FUNCTION_BLOCK MGE_Generico (* Multimedidor PM5300 - HidrycoLib *)
  (* Standard: 61499-2 *)
  (* Version 1.5, 15/10/2026, Hidryco, Hidryco, 1.5: tags de valores do IThis com prefixo STS_ (STS_TENSAO_*, STS_CORRENTE_*, STS_POTENCIA_*, STS_FATOR_POTENCIAL_TOTAL, STS_FREQUENCIA). 1.4: corrente A, B e C baixa (STP_CORRENTE_L, 3 alarmes, retardo STP_TEMPO_CORRENTE). 1.3: so as grandezas, ajustes e alarmes da especificacao do cliente (tensoes AB/BC/CA/AN/BN/CN, correntes A/B/C, potencias ativa e reativa A/B/C/total, frequencia, FP e aparente total; alarmes de comunicacao, FP baixo, tensao FF/FN alta/baixa, corrente A/B/C alta e frequencia alta/baixa). Referencia 0 = alarme desligado; um tempo de retardo por grupo. Os grupos de symlink continuam assinando tudo o que o PM53xxMbtcp publica, mas so as grandezas da especificacao entram na logica. 1.2: alarmes conforme a lista do cliente - falta de fase, tensao FF alta/baixa, tensao FN alta/baixa, corrente A/B/C alta, FP baixo, frequencia alta/baixa e falha de comunicacao (sai a corrente L). 1.1: Frequency do PM53xxMbtcp e VTQLINT: stsFrequencia passa para o grupo das energias (VTQLINT). 1.0: multimedidor PowerLogic PM5300 lido pelo HW CAT SE.FieldDevice.PM53xxMbtcp. Os symlinks do HW CAT (VTQREAL/VTQLINT) apontam para ${PATH}stsTensaoAB ... ${PATH}stsEnergiaAparente e ${PATH}stsComunicacaoOK/stsConexao/stsConexaoInt. Falta de fase, tensao H/L e corrente H/L ajustaveis na IHM (memorizados ate o reset). Tags do IThis com os nomes do CAT MGE antigo. *)
  PACKAGE Hidryco.HidrycoLib;
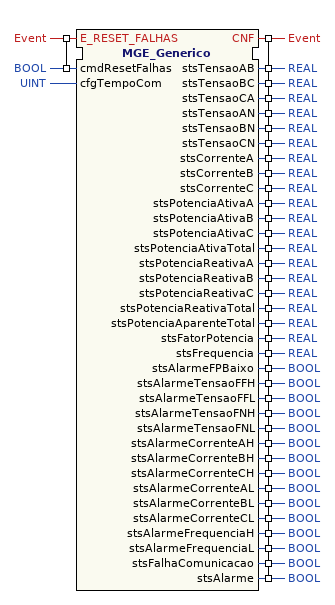
  EVENT_INPUT
    E_RESET_FALHAS WITH cmdResetFalhas; (* Reset pelo processo com cmdResetFalhas = TRUE *)
  END_EVENT
  EVENT_OUTPUT
    CNF WITH stsTensaoAB, stsTensaoBC, stsTensaoCA, stsTensaoAN, stsTensaoBN, stsTensaoCN, stsCorrenteA, stsCorrenteB, stsCorrenteC, stsPotenciaAtivaA, stsPotenciaAtivaB, stsPotenciaAtivaC, stsPotenciaAtivaTotal, stsPotenciaReativaA, stsPotenciaReativaB, stsPotenciaReativaC, stsPotenciaReativaTotal, stsPotenciaAparenteTotal, stsFatorPotencia, stsFrequencia, stsAlarmeFPBaixo, stsAlarmeTensaoFFH, stsAlarmeTensaoFFL, stsAlarmeTensaoFNH, stsAlarmeTensaoFNL, stsAlarmeCorrenteAH, stsAlarmeCorrenteBH, stsAlarmeCorrenteCH, stsAlarmeCorrenteAL, stsAlarmeCorrenteBL, stsAlarmeCorrenteCL, stsAlarmeFrequenciaH, stsAlarmeFrequenciaL, stsFalhaComunicacao, stsAlarme; (* Valores e alarmes (so na mudanca) *)
  END_EVENT
  VAR_INPUT
    cmdResetFalhas : BOOL; (* TRUE = reset (com o evento E_RESET_FALHAS) *)
    cfgTempoCom : UINT := 5; (* Tempo (s) sem comunicacao com o medidor para confirmar a falha *)
  END_VAR
  VAR_OUTPUT
    stsTensaoAB : REAL; (* Tensao A-B (V) *)
    stsTensaoBC : REAL; (* Tensao B-C (V) *)
    stsTensaoCA : REAL; (* Tensao C-A (V) *)
    stsTensaoAN : REAL; (* Tensao A-N (V) *)
    stsTensaoBN : REAL; (* Tensao B-N (V) *)
    stsTensaoCN : REAL; (* Tensao C-N (V) *)
    stsCorrenteA : REAL; (* Corrente fase A (A) *)
    stsCorrenteB : REAL; (* Corrente fase B (A) *)
    stsCorrenteC : REAL; (* Corrente fase C (A) *)
    stsPotenciaAtivaA : REAL; (* Potencia ativa fase A (kW) *)
    stsPotenciaAtivaB : REAL; (* Potencia ativa fase B (kW) *)
    stsPotenciaAtivaC : REAL; (* Potencia ativa fase C (kW) *)
    stsPotenciaAtivaTotal : REAL; (* Potencia ativa total (kW) *)
    stsPotenciaReativaA : REAL; (* Potencia reativa fase A (kVAr) *)
    stsPotenciaReativaB : REAL; (* Potencia reativa fase B (kVAr) *)
    stsPotenciaReativaC : REAL; (* Potencia reativa fase C (kVAr) *)
    stsPotenciaReativaTotal : REAL; (* Potencia reativa total (kVAr) *)
    stsPotenciaAparenteTotal : REAL; (* Potencia aparente total (kVA) *)
    stsFatorPotencia : REAL; (* Fator de potencia total *)
    stsFrequencia : REAL; (* Frequencia (Hz) *)
    stsAlarmeFPBaixo : BOOL; (* Fator de potência baixo (memorizado ate o reconhecimento) *)
    stsAlarmeTensaoFFH : BOOL; (* Tensão entre fases alta (memorizado ate o reconhecimento) *)
    stsAlarmeTensaoFFL : BOOL; (* Tensão entre fases baixa (memorizado ate o reconhecimento) *)
    stsAlarmeTensaoFNH : BOOL; (* Tensão fase-neutro alta (memorizado ate o reconhecimento) *)
    stsAlarmeTensaoFNL : BOOL; (* Tensão fase-neutro baixa (memorizado ate o reconhecimento) *)
    stsAlarmeCorrenteAH : BOOL; (* Corrente fase A alta (memorizado ate o reconhecimento) *)
    stsAlarmeCorrenteBH : BOOL; (* Corrente fase B alta (memorizado ate o reconhecimento) *)
    stsAlarmeCorrenteCH : BOOL; (* Corrente fase C alta (memorizado ate o reconhecimento) *)
    stsAlarmeCorrenteAL : BOOL; (* Corrente fase A baixa (memorizado ate o reconhecimento) *)
    stsAlarmeCorrenteBL : BOOL; (* Corrente fase B baixa (memorizado ate o reconhecimento) *)
    stsAlarmeCorrenteCL : BOOL; (* Corrente fase C baixa (memorizado ate o reconhecimento) *)
    stsAlarmeFrequenciaH : BOOL; (* Frequência alta (memorizado ate o reconhecimento) *)
    stsAlarmeFrequenciaL : BOOL; (* Frequência baixa (memorizado ate o reconhecimento) *)
    stsFalhaComunicacao : BOOL; (* Falha de comunicacao com o medidor *)
    stsAlarme : BOOL; (* Algum alarme do medidor *)
  END_VAR
  FBS
    IThis : MGE_Generico_HMI(QI := TRUE);
    plcStart1 : plcStart(Prio := 10);
    Logica : basicMGEGenerico;
    Tick : E_CYCLE(DT := T#1s);
    Tensoes : SYMLINKMULTIVARDST_2295B2715D3FE1C95(NAME1 := '$${PATH}stsTensaoAB', NAME2 := '$${PATH}stsTensaoBC', NAME3 := '$${PATH}stsTensaoCA', NAME4 := '$${PATH}stsTensaoMediaLL', NAME5 := '$${PATH}stsTensaoAN', NAME6 := '$${PATH}stsTensaoBN', NAME7 := '$${PATH}stsTensaoCN', NAME8 := '$${PATH}stsTensaoMediaLN', NAME9 := '$${PATH}stsDesequilibrioTensao', QI := TRUE); {SET_ATTRIBUTE(Configuration.GenericFBType.InterfaceParams, Runtime.System#I:=9;VALUE${I$}:VTQREAL,VTQREAL,VTQREAL,VTQREAL,VTQREAL,VTQREAL,VTQREAL,VTQREAL,VTQREAL)}
    Correntes : SYMLINKMULTIVARDST_858FA8D101163416(NAME1 := '$${PATH}stsCorrenteA', NAME2 := '$${PATH}stsCorrenteB', NAME3 := '$${PATH}stsCorrenteC', NAME4 := '$${PATH}stsCorrenteMedia', QI := TRUE); {SET_ATTRIBUTE(Configuration.GenericFBType.InterfaceParams, Runtime.System#I:=4;VALUE${I$}:VTQREAL,VTQREAL,VTQREAL,VTQREAL)}
    Potencias : SYMLINKMULTIVARDST_35CF2AFB1BB2205F(NAME1 := '$${PATH}stsPotenciaAtivaA', NAME2 := '$${PATH}stsPotenciaAtivaB', NAME3 := '$${PATH}stsPotenciaAtivaC', NAME4 := '$${PATH}stsPotenciaAtivaTotal', NAME5 := '$${PATH}stsPotenciaReativaA', NAME6 := '$${PATH}stsPotenciaReativaB', NAME7 := '$${PATH}stsPotenciaReativaC', NAME8 := '$${PATH}stsPotenciaReativaTotal', NAME9 := '$${PATH}stsPotenciaAparenteA', NAME10 := '$${PATH}stsPotenciaAparenteB', NAME11 := '$${PATH}stsPotenciaAparenteC', NAME12 := '$${PATH}stsPotenciaAparenteTotal', NAME13 := '$${PATH}stsFatorPotencia', QI := TRUE); {SET_ATTRIBUTE(Configuration.GenericFBType.InterfaceParams, Runtime.System#I:=13;VALUE${I$}:VTQREAL,VTQREAL,VTQREAL,VTQREAL,VTQREAL,VTQREAL,VTQREAL,VTQREAL,VTQREAL,VTQREAL,VTQREAL,VTQREAL,VTQREAL)}
    Energias : SYMLINKMULTIVARDST_9881907271BA9D7F(NAME1 := '$${PATH}stsEnergiaAtiva', NAME2 := '$${PATH}stsEnergiaReativa', NAME3 := '$${PATH}stsEnergiaAparente', NAME4 := '$${PATH}stsFrequencia', QI := TRUE); {SET_ATTRIBUTE(Configuration.GenericFBType.InterfaceParams, Runtime.System#I:=4;VALUE${I$}:VTQLINT,VTQLINT,VTQLINT,VTQLINT)}
    Comunicacao : SYMLINKMULTIVARDST_10236CFCCF63A5DF(NAME1 := '$${PATH}stsComunicacaoOK', NAME2 := '$${PATH}stsConexao', NAME3 := '$${PATH}stsConexaoInt', QI := TRUE); {SET_ATTRIBUTE(Configuration.GenericFBType.InterfaceParams, Runtime.System#I:=3;VALUE${I$}:BOOL,STRING,INT)}
    AlarmeFPL : ALARM_BIT(TYPE := 1, ACKTYPE_1 := 2, ACTIVE := TRUE); {SET_ATTRIBUTE(HMI.AlarmText, Fator de potência baixo)} {SET_ATTRIBUTE(HMI.AlarmClass, Warning)}
    AlarmeVFH : ALARM_BIT(TYPE := 1, ACKTYPE_1 := 2, ACTIVE := TRUE); {SET_ATTRIBUTE(HMI.AlarmText, Tensão entre fases alta)} {SET_ATTRIBUTE(HMI.AlarmClass, Warning)}
    AlarmeVFL : ALARM_BIT(TYPE := 1, ACKTYPE_1 := 2, ACTIVE := TRUE); {SET_ATTRIBUTE(HMI.AlarmText, Tensão entre fases baixa)} {SET_ATTRIBUTE(HMI.AlarmClass, Warning)}
    AlarmeVNH : ALARM_BIT(TYPE := 1, ACKTYPE_1 := 2, ACTIVE := TRUE); {SET_ATTRIBUTE(HMI.AlarmText, Tensão fase-neutro alta)} {SET_ATTRIBUTE(HMI.AlarmClass, Warning)}
    AlarmeVNL : ALARM_BIT(TYPE := 1, ACKTYPE_1 := 2, ACTIVE := TRUE); {SET_ATTRIBUTE(HMI.AlarmText, Tensão fase-neutro baixa)} {SET_ATTRIBUTE(HMI.AlarmClass, Warning)}
    AlarmeIAH : ALARM_BIT(TYPE := 1, ACKTYPE_1 := 2, ACTIVE := TRUE); {SET_ATTRIBUTE(HMI.AlarmText, Corrente da fase A alta)} {SET_ATTRIBUTE(HMI.AlarmClass, Warning)}
    AlarmeIBH : ALARM_BIT(TYPE := 1, ACKTYPE_1 := 2, ACTIVE := TRUE); {SET_ATTRIBUTE(HMI.AlarmText, Corrente da fase B alta)} {SET_ATTRIBUTE(HMI.AlarmClass, Warning)}
    AlarmeICH : ALARM_BIT(TYPE := 1, ACKTYPE_1 := 2, ACTIVE := TRUE); {SET_ATTRIBUTE(HMI.AlarmText, Corrente da fase C alta)} {SET_ATTRIBUTE(HMI.AlarmClass, Warning)}
    AlarmeIAL : ALARM_BIT(TYPE := 1, ACKTYPE_1 := 2, ACTIVE := TRUE); {SET_ATTRIBUTE(HMI.AlarmText, Corrente da fase A baixa)} {SET_ATTRIBUTE(HMI.AlarmClass, Warning)}
    AlarmeIBL : ALARM_BIT(TYPE := 1, ACKTYPE_1 := 2, ACTIVE := TRUE); {SET_ATTRIBUTE(HMI.AlarmText, Corrente da fase B baixa)} {SET_ATTRIBUTE(HMI.AlarmClass, Warning)}
    AlarmeICL : ALARM_BIT(TYPE := 1, ACKTYPE_1 := 2, ACTIVE := TRUE); {SET_ATTRIBUTE(HMI.AlarmText, Corrente da fase C baixa)} {SET_ATTRIBUTE(HMI.AlarmClass, Warning)}
    AlarmeFRH : ALARM_BIT(TYPE := 1, ACKTYPE_1 := 2, ACTIVE := TRUE); {SET_ATTRIBUTE(HMI.AlarmText, Frequência alta)} {SET_ATTRIBUTE(HMI.AlarmClass, Warning)}
    AlarmeFRL : ALARM_BIT(TYPE := 1, ACKTYPE_1 := 2, ACTIVE := TRUE); {SET_ATTRIBUTE(HMI.AlarmText, Frequência baixa)} {SET_ATTRIBUTE(HMI.AlarmClass, Warning)}
    AlarmeComunicacao : ALARM_BIT(TYPE := 1, ACKTYPE_1 := 2, ACTIVE := TRUE); {SET_ATTRIBUTE(HMI.AlarmText, Multimedidor sem comunicação)}
  END_FBS
  EVENT_CONNECTIONS
    plcStart1.FIRST_INIT TO IThis.A90CA12D67019FB2;
    plcStart1.REDO_INIT TO IThis.A90CA12D67019FB2;
    IThis.DF3130DED214D9B5 TO Logica.9F5D02D43587CE34;
    Logica.E47EE255A9E81DEF TO Tick.START;
    Logica.E47EE255A9E81DEF TO Tensoes.INIT;
    Logica.E47EE255A9E81DEF TO Correntes.INIT;
    Logica.E47EE255A9E81DEF TO Potencias.INIT;
    Logica.E47EE255A9E81DEF TO Energias.INIT;
    Logica.E47EE255A9E81DEF TO Comunicacao.INIT;
    Logica.E47EE255A9E81DEF TO AlarmeFPL.INIT;
    AlarmeFPL.INITO TO AlarmeFPL.REQ_INITDATA;
    AlarmeFPL.CNF_INITDATA TO AlarmeFPL.ACTIVATE;
    AlarmeFPL.INITO TO AlarmeVFH.INIT;
    AlarmeVFH.INITO TO AlarmeVFH.REQ_INITDATA;
    AlarmeVFH.CNF_INITDATA TO AlarmeVFH.ACTIVATE;
    AlarmeVFH.INITO TO AlarmeVFL.INIT;
    AlarmeVFL.INITO TO AlarmeVFL.REQ_INITDATA;
    AlarmeVFL.CNF_INITDATA TO AlarmeVFL.ACTIVATE;
    AlarmeVFL.INITO TO AlarmeVNH.INIT;
    AlarmeVNH.INITO TO AlarmeVNH.REQ_INITDATA;
    AlarmeVNH.CNF_INITDATA TO AlarmeVNH.ACTIVATE;
    AlarmeVNH.INITO TO AlarmeVNL.INIT;
    AlarmeVNL.INITO TO AlarmeVNL.REQ_INITDATA;
    AlarmeVNL.CNF_INITDATA TO AlarmeVNL.ACTIVATE;
    AlarmeVNL.INITO TO AlarmeIAH.INIT;
    AlarmeIAH.INITO TO AlarmeIAH.REQ_INITDATA;
    AlarmeIAH.CNF_INITDATA TO AlarmeIAH.ACTIVATE;
    AlarmeIAH.INITO TO AlarmeIBH.INIT;
    AlarmeIBH.INITO TO AlarmeIBH.REQ_INITDATA;
    AlarmeIBH.CNF_INITDATA TO AlarmeIBH.ACTIVATE;
    AlarmeIBH.INITO TO AlarmeICH.INIT;
    AlarmeICH.INITO TO AlarmeICH.REQ_INITDATA;
    AlarmeICH.CNF_INITDATA TO AlarmeICH.ACTIVATE;
    AlarmeICH.INITO TO AlarmeIAL.INIT;
    AlarmeIAL.INITO TO AlarmeIAL.REQ_INITDATA;
    AlarmeIAL.CNF_INITDATA TO AlarmeIAL.ACTIVATE;
    AlarmeIAL.INITO TO AlarmeIBL.INIT;
    AlarmeIBL.INITO TO AlarmeIBL.REQ_INITDATA;
    AlarmeIBL.CNF_INITDATA TO AlarmeIBL.ACTIVATE;
    AlarmeIBL.INITO TO AlarmeICL.INIT;
    AlarmeICL.INITO TO AlarmeICL.REQ_INITDATA;
    AlarmeICL.CNF_INITDATA TO AlarmeICL.ACTIVATE;
    AlarmeICL.INITO TO AlarmeFRH.INIT;
    AlarmeFRH.INITO TO AlarmeFRH.REQ_INITDATA;
    AlarmeFRH.CNF_INITDATA TO AlarmeFRH.ACTIVATE;
    AlarmeFRH.INITO TO AlarmeFRL.INIT;
    AlarmeFRL.INITO TO AlarmeFRL.REQ_INITDATA;
    AlarmeFRL.CNF_INITDATA TO AlarmeFRL.ACTIVATE;
    AlarmeFRL.INITO TO AlarmeComunicacao.INIT;
    AlarmeComunicacao.INITO TO AlarmeComunicacao.REQ_INITDATA;
    AlarmeComunicacao.CNF_INITDATA TO AlarmeComunicacao.ACTIVATE;
    AlarmeComunicacao.INITO TO plcStart1.ACK_FIRST;
    AlarmeComunicacao.INITO TO IThis.C08AD0831FA58CED;
    IThis.5861B63F088ADBAD TO Logica.6A49606260A35652;
    IThis.3F31327172D85BDC TO Logica.A0F14ADAA28E4173;
    E_RESET_FALHAS TO Logica.DB1848E569BB8432;
    Tick.EO TO Logica.DF07E6CBFE092BB1;
    Logica.AEC7342932406D99 TO CNF;
    Logica.9B7481123393F975 TO IThis.00C6D36E07251F2F;
    Tensoes.CNF TO Logica.F5C71D3E4D52B580;
    Correntes.CNF TO Logica.967BB9475D5FB31F;
    Potencias.CNF TO Logica.74289281190DCCEA;
    Energias.CNF TO Logica.8C17181F30D9640C;
    Comunicacao.CNF TO Logica.2AA09F5D795E9774;
    Logica.CA7EE46F7F0770BC TO AlarmeFPL.REQ;
    Logica.CA7EE46F7F0770BC TO AlarmeVFH.REQ;
    Logica.CA7EE46F7F0770BC TO AlarmeVFL.REQ;
    Logica.CA7EE46F7F0770BC TO AlarmeVNH.REQ;
    Logica.CA7EE46F7F0770BC TO AlarmeVNL.REQ;
    Logica.CA7EE46F7F0770BC TO AlarmeIAH.REQ;
    Logica.CA7EE46F7F0770BC TO AlarmeIBH.REQ;
    Logica.CA7EE46F7F0770BC TO AlarmeICH.REQ;
    Logica.CA7EE46F7F0770BC TO AlarmeIAL.REQ;
    Logica.CA7EE46F7F0770BC TO AlarmeIBL.REQ;
    Logica.CA7EE46F7F0770BC TO AlarmeICL.REQ;
    Logica.CA7EE46F7F0770BC TO AlarmeFRH.REQ;
    Logica.CA7EE46F7F0770BC TO AlarmeFRL.REQ;
    Logica.CA7EE46F7F0770BC TO AlarmeComunicacao.REQ;
    AlarmeFPL.IND_1 TO IThis.00C6D36E07251F2F;
    AlarmeVFH.IND_1 TO IThis.00C6D36E07251F2F;
    AlarmeVFL.IND_1 TO IThis.00C6D36E07251F2F;
    AlarmeVNH.IND_1 TO IThis.00C6D36E07251F2F;
    AlarmeVNL.IND_1 TO IThis.00C6D36E07251F2F;
    AlarmeIAH.IND_1 TO IThis.00C6D36E07251F2F;
    AlarmeIBH.IND_1 TO IThis.00C6D36E07251F2F;
    AlarmeICH.IND_1 TO IThis.00C6D36E07251F2F;
    AlarmeIAL.IND_1 TO IThis.00C6D36E07251F2F;
    AlarmeIBL.IND_1 TO IThis.00C6D36E07251F2F;
    AlarmeICL.IND_1 TO IThis.00C6D36E07251F2F;
    AlarmeFRH.IND_1 TO IThis.00C6D36E07251F2F;
    AlarmeFRL.IND_1 TO IThis.00C6D36E07251F2F;
    AlarmeComunicacao.IND_1 TO IThis.00C6D36E07251F2F;
    IThis.3F31327172D85BDC TO AlarmeFPL.ACK_C1;
    IThis.3F31327172D85BDC TO AlarmeVFH.ACK_C1;
    IThis.3F31327172D85BDC TO AlarmeVFL.ACK_C1;
    IThis.3F31327172D85BDC TO AlarmeVNH.ACK_C1;
    IThis.3F31327172D85BDC TO AlarmeVNL.ACK_C1;
    IThis.3F31327172D85BDC TO AlarmeIAH.ACK_C1;
    IThis.3F31327172D85BDC TO AlarmeIBH.ACK_C1;
    IThis.3F31327172D85BDC TO AlarmeICH.ACK_C1;
    IThis.3F31327172D85BDC TO AlarmeIAL.ACK_C1;
    IThis.3F31327172D85BDC TO AlarmeIBL.ACK_C1;
    IThis.3F31327172D85BDC TO AlarmeICL.ACK_C1;
    IThis.3F31327172D85BDC TO AlarmeFRH.ACK_C1;
    IThis.3F31327172D85BDC TO AlarmeFRL.ACK_C1;
    IThis.3F31327172D85BDC TO AlarmeComunicacao.ACK_C1;
  END_CONNECTIONS
  DATA_CONNECTIONS
    cfgTempoCom TO Logica.437048CAB4EF459B;
    cmdResetFalhas TO Logica.742F5E7E634543E1;
    Tensoes.VALUE1 TO Logica.23895DD175C25514;
    Tensoes.VALUE2 TO Logica.F90E2B2FC55BA1CA;
    Tensoes.VALUE3 TO Logica.9A2FEDFAA23B9FBE;
    Tensoes.VALUE5 TO Logica.EA2CDED484FB370F;
    Tensoes.VALUE6 TO Logica.45C7F73083D33855;
    Tensoes.VALUE7 TO Logica.49C54F216B8FD3B5;
    Correntes.VALUE1 TO Logica.15EFB699F1661CF7;
    Correntes.VALUE2 TO Logica.8E04AD2CCA4792B9;
    Correntes.VALUE3 TO Logica.8A2E8DB094282CC1;
    Potencias.VALUE1 TO Logica.8279BBA83A66993B;
    Potencias.VALUE2 TO Logica.F3D3261550357656;
    Potencias.VALUE3 TO Logica.1521741E9F36758F;
    Potencias.VALUE4 TO Logica.13CE1AEB225E8F43;
    Potencias.VALUE5 TO Logica.31DEB4D01C782F4A;
    Potencias.VALUE6 TO Logica.D0DBE61D0296D28C;
    Potencias.VALUE7 TO Logica.F287CB8A9A2AB36E;
    Potencias.VALUE8 TO Logica.B3A13548EF928803;
    Potencias.VALUE12 TO Logica.D657F63BBA25F39C;
    Potencias.VALUE13 TO Logica.505EEA3B9A786B68;
    Energias.VALUE4 TO Logica.29299DC668CC3955;
    Comunicacao.VALUE1 TO Logica.7B142F22116367BE;
    IThis.E6D256AC6C3A594B TO Logica.54EB28BC84E7838A;
    IThis.D4A3B585C3EA4F35 TO Logica.E9A3EA6D590FEE37;
    IThis.8EE9C7DEC4964674 TO Logica.4C3B3E1EC499BB7D;
    IThis.0FFBF509B5DA63B5 TO Logica.B3A7D982A721D879;
    IThis.4206B9E211992D1C TO Logica.05000A39B08793CD;
    IThis.AF82DCF1856B3FD7 TO Logica.DD5578AD81C8F373;
    IThis.2264561FF2B7379A TO Logica.70F112F8F27AB7E4;
    IThis.0646871FA8E56815 TO Logica.31CBD62CE860DD48;
    IThis.1539E10236608850 TO Logica.84C7AFD3C570D0FF;
    IThis.A68017885C22D1E2 TO Logica.0FCB7D8BABE5842B;
    IThis.B97C65AD134BAB6C TO Logica.5B2734CC365FC416;
    IThis.D88477A341E65E4E TO Logica.F9E02D7CA7FE396D;
    IThis.E3BBFB0CBE61AFDE TO Logica.B8BF3F3AEC8BA46F;
    IThis.D9D2C38C7AE71F9F TO Logica.09700DEBF5EDB7C8;
    Logica.D4D80A135835A68F TO AlarmeFPL.INP;
    Logica.C84C8E8A4AFB6B52 TO AlarmeVFH.INP;
    Logica.F520262A71826272 TO AlarmeVFL.INP;
    Logica.4400E5A533140BA8 TO AlarmeVNH.INP;
    Logica.7376632FDF9503CB TO AlarmeVNL.INP;
    Logica.63B40D626752D741 TO AlarmeIAH.INP;
    Logica.BD23AC0B2C0651A2 TO AlarmeIBH.INP;
    Logica.E5351E94A6A3DACF TO AlarmeICH.INP;
    Logica.2B9B0D1856474FB9 TO AlarmeIAL.INP;
    Logica.831D174108141DB9 TO AlarmeIBL.INP;
    Logica.8D40306CC7CC316D TO AlarmeICL.INP;
    Logica.B03E175FA415310D TO AlarmeFRH.INP;
    Logica.07A0D7C059B80A32 TO AlarmeFRL.INP;
    Logica.2BE8F70940E7CC3C TO AlarmeComunicacao.INP;
    Logica.D7A00C30A6619D8D TO stsTensaoAB;
    Logica.146C9A11D5258D71 TO stsTensaoBC;
    Logica.5A35EDE710ED9E91 TO stsTensaoCA;
    Logica.995DA9785F33D214 TO stsTensaoAN;
    Logica.55FA9C016450C2DD TO stsTensaoBN;
    Logica.59CA0F9C04715A67 TO stsTensaoCN;
    Logica.ADAF9D7DD197D4FE TO stsCorrenteA;
    Logica.C5BFFF1259440D18 TO stsCorrenteB;
    Logica.F325E224D7D277DF TO stsCorrenteC;
    Logica.A24B7F06D8ED8FA9 TO stsPotenciaAtivaA;
    Logica.978433C32C86D8EF TO stsPotenciaAtivaB;
    Logica.7E870D56C81A157A TO stsPotenciaAtivaC;
    Logica.04AF7B43BB533B3C TO stsPotenciaAtivaTotal;
    Logica.FD51813619FC2FED TO stsPotenciaReativaA;
    Logica.09C86328D003AC65 TO stsPotenciaReativaB;
    Logica.04CC3B6B399BF634 TO stsPotenciaReativaC;
    Logica.6FF4BBF46CE7DF72 TO stsPotenciaReativaTotal;
    Logica.B730EC83BF36AEFA TO stsPotenciaAparenteTotal;
    Logica.06F5ACACA7BE6E27 TO stsFatorPotencia;
    Logica.E3BC683E446C49CD TO stsFrequencia;
    Logica.0E52D748FE28BEED TO stsAlarmeFPBaixo;
    Logica.57FC50EADAB387B2 TO stsAlarmeTensaoFFH;
    Logica.0279D732904DE4AB TO stsAlarmeTensaoFFL;
    Logica.159CBC17837FAB70 TO stsAlarmeTensaoFNH;
    Logica.7F1B1FD426FC73B7 TO stsAlarmeTensaoFNL;
    Logica.260E565CCC5723A9 TO stsAlarmeCorrenteAH;
    Logica.7CCF92D2E693E51A TO stsAlarmeCorrenteBH;
    Logica.D74518AA6577BDAD TO stsAlarmeCorrenteCH;
    Logica.6990D128AAB2F344 TO stsAlarmeCorrenteAL;
    Logica.422EAD019B977526 TO stsAlarmeCorrenteBL;
    Logica.E808F4099E0C778F TO stsAlarmeCorrenteCL;
    Logica.70016D0B1A1C6D1D TO stsAlarmeFrequenciaH;
    Logica.0411BA8A94954963 TO stsAlarmeFrequenciaL;
    Logica.CC58FAB70A34AB27 TO stsFalhaComunicacao;
    Logica.803BAB84502C5F25 TO stsAlarme;
    Logica.D7A00C30A6619D8D TO IThis.1D73A57805826119;
    Logica.146C9A11D5258D71 TO IThis.7FAD3386F1FB5C1A;
    Logica.5A35EDE710ED9E91 TO IThis.AF7E451FC9E84A36;
    Logica.995DA9785F33D214 TO IThis.60CA7E27ABA7E199;
    Logica.55FA9C016450C2DD TO IThis.4D557000F41038EE;
    Logica.59CA0F9C04715A67 TO IThis.D896CE61D4A0C11F;
    Logica.ADAF9D7DD197D4FE TO IThis.88253584363F87AD;
    Logica.C5BFFF1259440D18 TO IThis.CCC2547F435CB96E;
    Logica.F325E224D7D277DF TO IThis.1436107BE30C06E0;
    Logica.A24B7F06D8ED8FA9 TO IThis.5CC3954CCBEF0AFC;
    Logica.978433C32C86D8EF TO IThis.A5BB1387B58C0213;
    Logica.7E870D56C81A157A TO IThis.B93512D8EE3E0FBB;
    Logica.04AF7B43BB533B3C TO IThis.C8432BCB562564AD;
    Logica.FD51813619FC2FED TO IThis.94236822BEBDDE08;
    Logica.09C86328D003AC65 TO IThis.6E4A4A5246FDF814;
    Logica.04CC3B6B399BF634 TO IThis.33FAEC88790E42C1;
    Logica.6FF4BBF46CE7DF72 TO IThis.02E12685E7B0E13F;
    Logica.B730EC83BF36AEFA TO IThis.9AD5849EE95B93D6;
    Logica.06F5ACACA7BE6E27 TO IThis.7780A13A457D6132;
    Logica.E3BC683E446C49CD TO IThis.7400873EEFE449B5;
    Logica.0E52D748FE28BEED TO IThis.4654ABD361B3B681;
    Logica.57FC50EADAB387B2 TO IThis.D6EC0E60D58ED0C1;
    Logica.0279D732904DE4AB TO IThis.FD7A3CEE3AC1D79E;
    Logica.159CBC17837FAB70 TO IThis.921CFD04CCBC8417;
    Logica.7F1B1FD426FC73B7 TO IThis.615BADE0B3B06AE1;
    Logica.260E565CCC5723A9 TO IThis.CA925D2D4BF76C39;
    Logica.7CCF92D2E693E51A TO IThis.A5D9B0BAD507C29D;
    Logica.D74518AA6577BDAD TO IThis.89B5AF8CDD0338CF;
    Logica.6990D128AAB2F344 TO IThis.4612D1904495E17C;
    Logica.422EAD019B977526 TO IThis.2EFB87AC5E7985FF;
    Logica.E808F4099E0C778F TO IThis.80943CA34CECFDDB;
    Logica.70016D0B1A1C6D1D TO IThis.0DDD122B567699FA;
    Logica.0411BA8A94954963 TO IThis.E18F931791B5F31E;
    Logica.CC58FAB70A34AB27 TO IThis.B9ADC96E13F532BB;
    Logica.803BAB84502C5F25 TO IThis.4850D614D76FCA73;
    AlarmeFPL.STATE_1 TO IThis.FBDA6FE625AC78F6;
    AlarmeVFH.STATE_1 TO IThis.B6758909339C2F62;
    AlarmeVFL.STATE_1 TO IThis.6AE1605DFEB7FD1F;
    AlarmeVNH.STATE_1 TO IThis.37DC20F04F565B38;
    AlarmeVNL.STATE_1 TO IThis.C2CC757D9BDD8819;
    AlarmeIAH.STATE_1 TO IThis.A325BC62EADB0D8C;
    AlarmeIBH.STATE_1 TO IThis.B7D8C028DEDB4DFD;
    AlarmeICH.STATE_1 TO IThis.E445999A8E957193;
    AlarmeIAL.STATE_1 TO IThis.0D2645BFB4559CB1;
    AlarmeIBL.STATE_1 TO IThis.130E1473E7C6095A;
    AlarmeICL.STATE_1 TO IThis.097533B7E775C720;
    AlarmeFRH.STATE_1 TO IThis.F1E72D82FF4DDF80;
    AlarmeFRL.STATE_1 TO IThis.0D1E5BCB23F4B165;
    AlarmeComunicacao.STATE_1 TO IThis.EC7EBE5361F4D581;
  END_CONNECTIONS
END_FUNCTION_BLOCK
